// TIA Portal V19 export
DATA_BLOCK "MB_TCP_CLIENT"   // DB18
{ S7_Optimized_Access := 'FALSE'; DB_Accessible_From_OPC_UA := 'FALSE' }
// stored: DBAccessibleFromOPCUA false
   VAR
      MB_CONNECT : TCON_IP_v4;
   END_VAR
BEGIN
   MB_CONNECT.InterfaceId := 64;
   MB_CONNECT.ID := 1;
   MB_CONNECT.ConnectionType := 11;
   MB_CONNECT.ActiveEstablished := 1;
   MB_CONNECT.RemoteAddress.ADDR[1] := 192;
   MB_CONNECT.RemoteAddress.ADDR[2] := 168;
   MB_CONNECT.RemoteAddress.ADDR[3] := 0;
   MB_CONNECT.RemoteAddress.ADDR[4] := 60;
   MB_CONNECT.RemotePort := 502;
END_DATA_BLOCK
